Fanuc KAREL source: KS00028.KL

PROGRAM KS00028
%NOLOCKGROUP
TYPE
  REC_T = STRUCTURE
    VALUE: INTEGER
    FLAG: BOOLEAN
  ENDSTRUCTURE
VAR
  A: QUEUE_TYPE
  B: QUEUE_TYPE
  FLAG: BOOLEAN
  N: INTEGER
  STATUS: INTEGER
  PN: STRING[80]
  VN: STRING[80]
BEGIN
  PN = ''
  VN = 'A'
  SET_VAR(N, PN, VN, A, STATUS)
END KS00028
